(* IEC 61131-3 sources: plc-vscode/tests/st/test-ready/rusty/tests/lit/multi/extern_st_polymorphism, 2 files *)

(* ---- app.st ---- *)
// Redeclare interface so the compiler knows the shape
INTERFACE IGreeter
    METHOD greet
    END_METHOD
END_INTERFACE

// External declaration — the real implementation is in libpoly.so
{external}
FUNCTION_BLOCK FbA IMPLEMENTS IGreeter
VAR
    id : DINT;
END_VAR
    METHOD greet
    END_METHOD
END_FUNCTION_BLOCK

FUNCTION main
VAR
    inst : FbA;
    pInst : POINTER TO FbA;
    iface : IGreeter;
END_VAR
    inst.id := 7;
    pInst := ADR(inst);

    // Dynamic vtable dispatch
    pInst^.greet();

    // Interface dispatch (itable)
    iface := inst;
    iface.greet();
END_FUNCTION

(* ---- lib.st ---- *)
INTERFACE IGreeter
    METHOD greet
    END_METHOD
END_INTERFACE

FUNCTION_BLOCK FbA IMPLEMENTS IGreeter
VAR
    id : DINT;
END_VAR
    METHOD greet
        printf('FbA::greet (id=%d)$N', THIS^.id);
    END_METHOD
END_FUNCTION_BLOCK
